			IF pResultCheck <> 0 AND Result = 0 THEN
				Result := pResultCheck;
				codeposition := CONCAT(CONCAT(__POUNAME(),'() / '),__POSITION());
			END_IF;
		END_IF;
		IF pResultCheck = 0 THEN
			count_cycle := 0;
			REPEAT			
				SysFile.SysFileWrite(hFileCheck,ADR(stReSa),TO_UINT(LEN(stReSa)),ADR(pResultCheck));
				count_cycle := count_cycle + 1;
			UNTIL
				pResultCheck = 0 OR count_cycle >= 100 
			END_REPEAT;						
		ELSE
			proError := TRUE;	
			IF Result = 0 THEN
				Result := 16#C7A;
				codeposition := CONCAT(CONCAT(__POUNAME(),'() / '),__POSITION());
			END_IF
		END_IF;  
	END_IF;  
END_IF;
END_METHOD

PROPERTY proFilePathCheckFile : STRING[255];
GET
// FILE Path auf SPS
 proFilePathCheckFile:= CONCAT(  
						CONCAT(  
						CONCAT(                                  
								'$$PlcLogic$$/',  
								'ConfigFiles/Actual/'),  
								stCodeDir),  
								'_Check.txt');
END_GET
END_PROPERTY

METHOD metChild
VAR_INPUT
	itfDataTypeObj  :   ITF_DATATYPE;
END_VAR
IF scState.xGetChild THEN
	IF __QUERYINTERFACE(itfDataTypeObj,itfDataTypeObj) THEN
		IF NOT itfDataTypeObj.proChildAddDone THEN
			usiLastChild := itfDataTypeObj.proparaNr;
			itfDataTypeObj.proChildAddDone := TRUE;
		END_IF;
	END_IF;
END_IF;
END_METHOD

{attribute 'monitoring':='call'}
PROPERTY proLoad : BOOL
GET
proLoad := GVL_Config.xLoad;
END_GET
END_PROPERTY

METHOD FINAL metSaveFile : BOOL
VAR_INPUT  
    itfDataTypeObj  :   ITF_DATATYPE;
END_VAR
VAR
    udiPos  : UDINT;
    stSave  : STRING[172];
	pulPos  : __XWORD;
    dwWrite : DWORD;
	saefty_count	:USINT;
END_VAR
IF hFile <> 0 AND pResult = 0 AND itfDataTypeObj.proParaNr > 0 THEN
    udiPos := LIMIT(1,itfDataTypeObj.proParaNr,255);
   IF udiPos = 1 THEN
        udiPos :=  0;  
        stSave := CONCAT(itfDataTypeObj.proStrPara,'$R'); 
    ELSE
        udiPos := (udiPos * GlobalKonstant.diLineSize) - GlobalKonstant.diLineSize -1;
        stSave := CONCAT('$N',CONCAT(itfDataTypeObj.proStrPara,'$R')); 
	END_IF;
	saefty_count	:= 0;
	REPEAT	
		pResult := SysFile.SysFileSetPos(hFile,0);
		pResult := SysFile.SysFileGetPos(hFile,ADR(pulPos));
		saefty_count := saefty_count + 1;
	UNTIL
		pResult = 0 OR saefty_count >= 10		
	END_REPEAT
	IF pResult <> 0 AND Result = 0 THEN
		Result := pResult;
		codeposition :=   CONCAT(CONCAT(CONCAT(CONCAT(CONCAT(CONCAT(__POUNAME(),'() / '),__POSITION()),' POSW= '),TO_STRING(udiPos)),' POSR='),TO_STRING(pulPos));
		status := SysFile.SysFileGetStatus(hFile);
	END_IF;
	IF pulPos <> udiPos THEN
		saefty_count	:= 0;
		REPEAT
			SysFile.SysFileFlush(hFile);
			pResult := SysFile.SysFileSetPos(hFile,udiPos);
			saefty_count := saefty_count + 1;
		UNTIL
			pResult = 0 OR saefty_count >= 10		
		END_REPEAT
	END_IF;
	IF pResult <> 0 AND Result = 0 THEN
		Result := pResult;
		codeposition :=   CONCAT(CONCAT(CONCAT(CONCAT(CONCAT(CONCAT(__POUNAME(),'() / '),__POSITION()),' POSW= '),TO_STRING(udiPos)),' POSR='),TO_STRING(pulPos));
	END_IF;
    IF hFile <> 0 AND pResult = 0 THEN
		REPEAT 
			pResult := SysFile.SysFileSetPos(hFile,udiPos);
			dwWrite := TO_DWORD(SysFile.SysFileWrite(hFile,ADR(stSave),TO_UDINT(LEN(stSave)),ADR(pResult)));
			SysFile.SysFileFlush(hFile);
			saefty_count := saefty_count + 1;
		UNTIL
			pResult = 0 OR saefty_count >= 10	
		END_REPEAT
		IF pResult <> 0 AND Result = 0 THEN
			Result := pResult;
			codeposition := CONCAT(CONCAT(__POUNAME(),'() / '),__POSITION());
			status := SysFile.SysFileGetStatus(hFile);
		END_IF;
    END_IF;
END_IF;
IF pResult <> 0 THEN
    pResult := pResult;
ELSE
    metSaveFile := NOT TO_BOOL(pResult) AND dwWrite = TO_UDINT(LEN(stSave));
END_IF
scState.xEventSave := TRUE;
END_METHOD

METHOD FINAL metSave : BOOL
VAR_INPUT
    itfDataTypeObj  :   ITF_DATATYPE;
END_VAR
VAR
    uiSafetyCount   :   UINT;
    wPos            :   WORD;
    xSysSemapohre   :   BOOL;
END_VAR
IF proSave OR itfDataTypeObj.proSaveOnChange THEN  
    IF NOT itfDataTypeObj.proIsSaving THEN 
        itfDataTypeObj.proIsSaving := TRUE;
        xSysSemapohre := TRUE;   
    END_IF;
    IF xSysSemapohre THEN
        uiSafetyCount := 0;           
        REPEAT
            pResult := 0; 
            (* File Lesen *)
            IF NOT scState.xIsOpen THEN
                scState.xIsOpen := metOpenFile();
            END_IF;    
            IF scState.xIsOpen THEN
                metSave := metSaveFile(itfDataTypeObj);  
            END_IF;
            uiSafetyCount := uiSafetyCount + 1;
        UNTIL
            metSave = TRUE OR uiSafetyCount = 16#000F
        END_REPEAT
        IF NOT metSave THEN
            THIS^.proError      := TRUE;
            THIS^.proErrorNr    := itfDataTypeObj.proParaNr;
			IF Result = 0 THEN
				Result := 16#C7A;
				codeposition := CONCAT(CONCAT(__POUNAME(),'() / '),__POSITION());
			END_IF
        END_IF  
        xSysSemapohre := FALSE;
        itfDataTypeObj.proIsSaving      := FALSE;
        itfDataTypeObj.proSaveOnChange  := FALSE;		
    END_IF;
END_IF;
END_METHOD

PROPERTY proError : BOOL
GET
proError := xError;
END_GET
SET
xError := proError;
END_SET
END_PROPERTY

{attribute 'monitoring_encoding' := 'UTF-8'}
PROPERTY proFilePath : STRING[255];
GET
// FILE Path auf SPS
proFilePath	     :=      	CONCAT(
							CONCAT(
							CONCAT(                                
									'$$PlcLogic$$/',
									'ConfigFiles/Actual/'),
									stCodeDir),
									'_Config.txt');                                  
								
IF proLoad OR proSave THEN
	proFilePath	    :=      CONCAT(
							CONCAT(
							CONCAT(    
							CONCAT(                            
									'$$PlcLogic$$/',
									'ConfigFiles/'),
									GVL_Config.stBackUp),
									stCodeDir),
									'_Config.txt');  
END_IF;
END_GET
END_PROPERTY

METHOD metCleanUpInit
VAR_INPUT
END_VAR
pResult     		:= fcFileClose(hFile,stCodeDir,'FbConfigFile CleanupIni Z1');
hFile       		:= SysTypes.RTS_INVALID_HANDLE;
pResultCheck		:= fcFileClose(hFileCheck,stCodeDir,'FbConfigFile CleanupIni Z3');
hFileCheck  		:= SysTypes.RTS_INVALID_HANDLE;
fcFileDelete(proFilePathCheckFile);
scState.xInit       := FALSE;
scState.xInitDone	:= TRUE;
iCaseInit   		:= iCaseInit + 1;

IF pResult <> 0 AND Result = 0 THEN
	Result := pResult;
	codeposition := CONCAT(CONCAT(__POUNAME(),'() / '),__POSITION());
END_IF;
IF pResultCheck <> 0 AND Result = 0 THEN
	Result := pResultCheck;
	codeposition := CONCAT(CONCAT(__POUNAME(),'() / '),__POSITION());
END_IF;
END_METHOD

METHOD FINAL metInit : BOOL
VAR_INPUT
    itfDataTypeObj  :   ITF_DATATYPE;
END_VAR
IF scstate.xGetChild THEN
	metChild(itfDataTypeObj);
END_IF;
IF scState.xInit THEN
    IF metCheckNr(itfDataTypeObj,TRUE,FALSE) THEN
        IF NOT metLoadFile(itfDataTypeObj) THEN
            metSaveFile(itfDataTypeObj);
        END_IF;  
        metCheckNr(itfDataTypeObj,FALSE,TRUE);
		metInit := TRUE;
    ELSE    
        proError    := TRUE;
        proErrorNr  := itfDataTypeObj.proParaNr;        
		IF Result = 0 THEN
			Result := 16#C7A;
			codeposition := CONCAT(CONCAT(__POUNAME(),'() / '),__POSITION());
		END_IF
    END_IF;
	IF __QUERYINTERFACE(itfDataTypeObj,itfDataTypeObj) THEN
		IF itfDataTypeObj.proparaNr = usilastChild THEN
			metCleanUpInit();
		END_IF
	END_IF;         
END_IF;
END_METHOD

//FB_Init ist immer implizit verfügbar und wird primär für die Initialisierung verwendet.
//Der Rückgabewert wird nicht ausgewertet. Für gezielte Einflussnahme können Sie
//die Methoden explizit deklarieren und darin mit dem Standard-Initialisierungscode 
//zusätzlichen Code bereitstellen. Sie können den Rückgabewert auswerten.
METHOD FINAL FB_Init: BOOL
VAR_INPUT    
bInitRetains: BOOL; // TRUE: Die Retain-Variablen werden initialisiert (Reset warm / Reset kalt)    
bInCopyCode: BOOL;  // TRUE: Die Instanz wird danach in den Kopiercode kopiert (Online-Change)
END_VAR
hFile   := SysTypes.RTS_INVALID_HANDLE;
hFileCheck  := SysTypes.RTS_INVALID_HANDLE;
END_METHOD

{attribute 'monitoring':='call'}
PROPERTY proSave : BOOL
GET
proSave := GVL_Config.xSave;
END_GET
END_PROPERTY

{attribute 'monitoring':='call'}
PROPERTY proInitDone : BOOL
GET
proInitDone := scState.xInitDone;
END_GET
END_PROPERTY

PROPERTY ProSetInstancePathOnDynCreate : STRING(255)
SET
stCodeDir := ProSetInstancePathOnDynCreate;
metCodeDirCreate();
END_SET
END_PROPERTY

METHOD metCleanUp
VAR_INPUT	
END_VAR
pResult     		:= fcFileClose(hFile,stCodeDir,'FbConfigFile Cleanup Z1');
hFile       		:= SysTypes.RTS_INVALID_HANDLE;
scState.xIsOpen 	:= FALSE;
END_METHOD

METHOD metCheckLastChild
VAR_INPUT  
    itfDataTypeObj  :   ITF_DATATYPE;
END_VAR
IF __QUERYINTERFACE(itfDataTypeObj,itfDataTypeObj) THEN
	IF itfDataTypeObj.proparaNr = usilastChild THEN
		metCleanUp();
	END_IF
END_IF;
END_METHOD

END_FUNCTION_BLOCK

// 30 Program Organization Units/Basis/fbConfigFile
{attribute 'enable_dynamic_creation'}
{attribute 'hide_all_locals'}
{attribute 'reflection'} 
FUNCTION_BLOCK fbConfigFile IMPLEMENTS ITF_CONFIGFILE
VAR_OUTPUT
    xError              :   BOOL;
    uiErrorNr           :   UINT;
	Result              :   RTS_IEC_RESULT;
	codeposition		:	STRING(255);
	status					:	SysFile.SYS_FILE_STATUS;
END_VAR
VAR
    {attribute 'instance-path'} 
    {attribute 'noinit'}     
	{attribute 'monitoring_encoding' := 'UTF-8'}
    stCodeDir               :   STRING[255]; 
    iCaseInit               :   INT                 := 0;
    scState                 :   scStateConfigFile;
    hFile                   :   RTS_IEC_HANDLE;
    pResult                 :   RTS_IEC_RESULT;
    hFileCheck              :   RTS_IEC_HANDLE;
    pResultCheck            :   RTS_IEC_RESULT;    
	usiLastChild			:	USINT;
END_VAR

CASE iCaseInit OF
	0: // Get Last Child
		scState.xGetChild   := TRUE;
		metCodeDirCreate();
		iCaseInit := iCaseInit + 1;
	1: // Init
		scState.xGetChild	:= FALSE;
        scState.xInit       := TRUE;
		
		hFile := fcFileOpen(proFilePath,SysFile.ACCESS_MODE.AM_APPEND_PLUS,pResult);
		IF hFile <> SysTypes.RTS_INVALID_HANDLE THEN
			SysFile.SysFileSetPos(hFile,0);
		END_IF;
		// Check File
		hFileCheck := fcFileOpen(proFilePathCheckFile,SysFile.ACCESS_MODE.AM_WRITE_PLUS,pResultCheck);
		iCaseInit   := iCaseInit + 1;
	2: // Init Done
		;	// Wait on Clean up Init Call
	3: // Check if Save or Load 
		IF (GVL_Config.xSave OR GVL_Config.xLoad) AND_THEN hFile = SysTypes.RTS_INVALID_HANDLE THEN
            scState.xIsOpen := metOpenFile();  
		END_IF;
	ELSE
		iCaseInit   := 0;   
END_CASE;
// Meldung 
IF NOT scState.xEventLoad AND NOT scState.xEventSave AND scState.xEventDetekted THEN
	scState.xEventDetekted := FALSE; 
END_IF;
IF scState.xEventSave THEN
	scState.xEventDetekted := TRUE;
	scState.xEventSave 	   := FALSE;    
END_IF;    
IF scState.xEventLoad THEN
	scState.xEventDetekted := TRUE;
	scState.xEventLoad     := FALSE;    
END_IF; 
IF xError AND_THEN NOT GVL_Config.xError THEN
    GVL_Config.xError 			:= TRUE;
    GVL_Config.stPath			:= stCodeDir;
	GVL_Config.Result			:= Result;
	GVL_Config.codeposition 	:= codeposition;
	GVL_Config.status			:= status;
END_IF;

METHOD FINAL metLoad : BOOL
VAR_INPUT  
    itfDataTypeObj  :   ITF_DATATYPE;
END_VAR
VAR
    uiSafetyCount   :   UINT;
END_VAR
IF proLoad THEN
    REPEAT
        pResult       := 0;
        IF NOT scState.xIsOpen THEN
            scState.xIsOpen := metOpenFile();    
		END_IF
        IF scState.xIsOpen THEN
            metLoad       := metLoadFile(itfDataTypeObj);  
        END_IF;    
            uiSafetyCount := uiSafetyCount + 1;
    UNTIL
        metLoad = TRUE OR uiSafetyCount = 16#FFFF
    END_REPEAT;     
    IF NOT metLoad THEN
        THIS^.proError      := TRUE;
        THIS^.proErrorNr    := itfDataTypeObj.proParaNr;
    END_IF; 
END_IF;
END_METHOD

METHOD metOpenFile : BOOL
VAR_INPUT
END_VAR
hFile   := fcFileOpen(proFilePath,SysFile.ACCESS_MODE.AM_READ_PLUS,pResult);
IF pResult = 0 AND hFile <> SysTypes.RTS_INVALID_HANDLE THEN
    metOpenFile := TRUE;
ELSE
    metOpenFile := FALSE;
END_IF
END_METHOD

PROPERTY proErrorNr : UINT
SET
uiErrorNr := proErrorNr;
END_SET
GET
proErrorNr := uiErrorNr;
END_GET
END_PROPERTY

METHOD PRIVATE FINAL metCodeDirCreate : BOOL
VAR
    uiFor                   :   UINT;
END_VAR
// Instanzpfad des Funktionsbausteinens in Ordnerstrucktur wandeln
FOR uiFor := 0 TO SIZEOF(stCodeDir)-1 DO
    // Punkt . durch Slash / ersetzen
    IF stCodeDir[uiFor] = 46 THEN
        stCodeDir[uiFor] := 47;
    END_IF;            
END_FOR;
END_METHOD

//FB_Exit muss explizit implementiert werden. Wenn es eine Implementierung gibt, dann wird 
//die Methode aufgerufen, bevor die Steuerung den Code der Funktionsbaustein-Instanz entfernt
//(impliziter Aufruf. Der Rückgabewert wird nicht ausgewertet.
METHOD FINAL FB_Exit: BOOL
VAR_INPUT    
    bInCopyCode: BOOL;  // TRUE: Die Exit-Methode wird aufgerufen, um die Instanz zu verlassen, die hinterher kopiert wird Online-Change).  
END_VAR
pResult := SysFile.SysFileClose(hFile);
hFile   := SysTypes.RTS_INVALID_HANDLE;
SysFile.SysFileClose(hFileCheck);
hFileCheck  := SysTypes.RTS_INVALID_HANDLE;
fcFileDelete(proFilePathCheckFile);
END_METHOD

{attribute 'monitoring':='call'}
PROPERTY proSave : BOOL
GET
proSave := GVL_Config.xSave;
END_GET
END_PROPERTY

METHOD FINAL metLoadFile : BOOL
VAR_INPUT  
    itfDataTypeObj  :   ITF_DATATYPE;
END_VAR
VAR
    udiPos  : UDINT;
    stRead  : STRING[170];
    xValid  : BOOL;
END_VAR
IF hFile <> SysTypes.RTS_INVALID_HANDLE AND itfDataTypeObj.proParaNr > 0 THEN
    udiPos := LIMIT(1,itfDataTypeObj.proParaNr,255);
   IF udiPos = 1 THEN
        udiPos :=  udiPos -1;   
    ELSE 
        udiPos := (udiPos * GlobalKonstant.diLineSize) - GlobalKonstant.diLineSize;
	END_IF;
    pResult := SysFile.SysFileSetPos(hFile,udiPos);
END_IF;
IF pResult = 0 AND hFile <> SysTypes.RTS_INVALID_HANDLE THEN
    SysFile.SysFileRead(hFile,ADR(stRead),GlobalKonstant.diStringSize,ADR(pResult));
    stRead[170] := 0;
    IF itfDataTypeObj.proParaNr = TO_UINT(MID(stRead,5,2)) THEN
        itfDataTypeObj.proStrPara := stRead;
        xValid := TRUE;
	END_IF;
END_IF;
metLoadFile := NOT TO_BOOL(pResult) AND xValid;
scState.xEventLoad := TRUE;
END_METHOD

PROPERTY proEventDetekted : BOOL
GET
proEventDetekted := scState.xEventDetekted;
END_GET
END_PROPERTY

METHOD FINAL metCheckNr : BOOL
VAR_INPUT
    itfDataTypeObj  :   ITF_DATATYPE;
    xCheck          :   BOOL;
    xCheckDone      :   BOOL;
END_VAR
VAR
    udiPos  : UDINT;
    stReSa  : STRING[1];
    xValid  : BOOL;
    pulPos  : DWORD;
END_VAR
IF xCheck THEN
    IF pResultCheck = 0 AND itfDataTypeObj.proParaNr > 0 THEN
        udiPos := LIMIT(1,itfDataTypeObj.proParaNr,255)-1;
        pResultCheck := SysFile.SysFileSetPos(hFileCheck,udiPos);
	ELSE
		set_error(CONCAT(CONCAT(__POUNAME(),'() / '),__POSITION()),pResultCheck);
    END_IF;
    IF pResultCheck = 0 THEN
        SysFile.SysFileRead(hFileCheck,ADR(stReSa),1,ADR(pResultCheck));
        IF TO_INT(stReSa) = 1 THEN
            xValid 		:= FALSE; 
			proError 	:= TRUE;
			proErrorNr 	:= itfDataTypeObj.proParaNr;
        ELSE
            xValid := TRUE; 
		END_IF
	ELSE
		proError := TRUE;
		set_error(CONCAT(CONCAT(__POUNAME(),'() / '),__POSITION()),pResultCheck);
    END_IF;
    metCheckNr := NOT TO_BOOL(pResultCheck) AND xValid;
ELSIF xCheckDone THEN
    IF pResultCheck = 0 AND itfDataTypeObj.proParaNr > 0 THEN
            udiPos := LIMIT(1,itfDataTypeObj.proParaNr,255)-1;
            stReSa := TO_STRING(1);
            pResultCheck := SysFile.SysFileGetPos(hFileCheck,ADR(pulPos));
            pResultCheck := SysFile.SysFileSetPos(hFileCheck,udiPos);
            pResultCheck := SysFile.SysFileGetPos(hFileCheck,ADR(pulPos));
    END_IF;
    IF pResultCheck = 0 THEN
        SysFile.SysFileWrite(hFileCheck,ADR(stReSa),TO_UINT(LEN(stReSa)),ADR(pResultCheck));
	ELSE
		set_error(CONCAT(CONCAT(__POUNAME(),'() / '),__POSITION()),pResultCheck);
		proError := TRUE;	
    END_IF;    
END_IF;
END_METHOD

PROPERTY proFilePathCheckFile : STRING[255];
GET
// FILE Path auf SPS
 proFilePathCheckFile:= CONCAT(  
						CONCAT(  
						CONCAT(                                  
								'$$PlcLogic$$/',  
								'ConfigFiles/Actual/'),  
								stCodeDir),  
								'_Check.txt');
END_GET
END_PROPERTY

METHOD metChild
VAR_INPUT
	itfDataTypeObj  :   ITF_DATATYPE;
END_VAR
IF scState.xGetChild THEN
	IF __QUERYINTERFACE(itfDataTypeObj,itfDataTypeObj) THEN
		IF NOT itfDataTypeObj.proChildAddDone THEN
			usiLastChild := itfDataTypeObj.proparaNr;
			itfDataTypeObj.proChildAddDone := TRUE;
		END_IF;
	END_IF;
END_IF;
END_METHOD

PROPERTY proError : BOOL
GET
proError := xError;
END_GET
SET
xError := proError;
END_SET
END_PROPERTY

{attribute 'monitoring':='call'}
PROPERTY proLoad : BOOL
GET
proLoad := GVL_Config.xLoad;
END_GET
END_PROPERTY

METHOD FINAL metSaveFile : BOOL
VAR_INPUT  
    itfDataTypeObj  :   ITF_DATATYPE;
END_VAR
VAR
    udiPos  : UDINT;
    stSave  : STRING[172];
	pulPos  : DWORD;
    dwWrite : DWORD;
END_VAR
IF hFile <> SysTypes.RTS_INVALID_HANDLE AND pResult = 0 AND itfDataTypeObj.proParaNr > 0 THEN
    udiPos := LIMIT(1,itfDataTypeObj.proParaNr,255);
   IF udiPos = 1 THEN
        udiPos :=  udiPos -1;  
        stSave := CONCAT(itfDataTypeObj.proStrPara,'$R'); 
    ELSE
        udiPos := (udiPos * GlobalKonstant.diLineSize) - GlobalKonstant.diLineSize - 1;
        stSave := CONCAT('$N',CONCAT(itfDataTypeObj.proStrPara,'$R')); 
	END_IF;
        pResult := SysFile.SysFileGetPos(hFile,ADR(pulPos));
        pResult := SysFile.SysFileSetPos(hFile,udiPos);
        pResult := SysFile.SysFileGetPos(hFile,ADR(pulPos));
    IF hFile <> 0 AND pResult = 0 THEN
        dwWrite := TO_DWORD(SysFile.SysFileWrite(hFile,ADR(stSave),TO_UDINT(LEN(stSave)),ADR(pResult)));
	ELSE
		set_error(CONCAT(CONCAT(__POUNAME(),'() / '),__POSITION()),pResult);
    END_IF;
END_IF;
IF pResult <> 0 THEN
	set_error(CONCAT(CONCAT(__POUNAME(),'() / '),__POSITION()),pResult);
ELSE
    metSaveFile := NOT TO_BOOL(pResult) AND dwWrite = TO_UDINT(LEN(stSave));
END_IF
scState.xEventSave := TRUE;
END_METHOD

METHOD FINAL metSave : BOOL
VAR_INPUT
    itfDataTypeObj  :   ITF_DATATYPE;
END_VAR
VAR
    uiSafetyCount   :   UINT;
    wPos            :   WORD;
    xSysSemapohre   :   BOOL;
END_VAR
IF NOT xError THEN
	IF proSave OR itfDataTypeObj.proSaveOnChange THEN  
		IF NOT itfDataTypeObj.proIsSaving THEN 
			itfDataTypeObj.proIsSaving := TRUE;
			xSysSemapohre := TRUE;   
		END_IF;
		IF xSysSemapohre THEN
			uiSafetyCount := 0;           
			REPEAT
				pResult := 0; 
				(* File Lesen *)
				IF NOT scState.xIsOpen THEN
					scState.xIsOpen := metOpenFile();
				END_IF;    
				IF scState.xIsOpen THEN
					metSave := metSaveFile(itfDataTypeObj);  
				END_IF;
				uiSafetyCount := uiSafetyCount + 1;
				IF NOT metSave THEN
					wPos := 16#EEEE;    
				END_IF
			UNTIL
				metSave = TRUE OR uiSafetyCount = 16#FFFF
			END_REPEAT
			IF NOT metSave THEN
				THIS^.proError      := TRUE;
				THIS^.proErrorNr    := itfDataTypeObj.proParaNr;
			END_IF  
			xSysSemapohre := FALSE;
			itfDataTypeObj.proIsSaving      := FALSE;
			itfDataTypeObj.proSaveOnChange  := FALSE;		
		END_IF;
	END_IF;
END_IF;
END_METHOD

{attribute 'monitoring':='call'}
PROPERTY proInitDone : BOOL
GET
proInitDone := scState.xInitDone;
END_GET
END_PROPERTY

{attribute 'monitoring_encoding' := 'UTF-8'}
PROPERTY proFilePath : STRING[255];
GET
// FILE Path auf SPS
proFilePath     :=      	CONCAT(
							CONCAT(
							CONCAT(                                
									'$$PlcLogic$$/',
									'ConfigFiles/Actual/'),
									stCodeDir),
									'_Config.txt');                                  
								
IF proLoad OR proSave THEN
	proFilePath     :=      CONCAT(
							CONCAT(
							CONCAT(    
							CONCAT(                            
									'$$PlcLogic$$/',
									'ConfigFiles/'),
									GVL_Config.stBackUp),
									stCodeDir),
									'_Config.txt');  
END_IF;
END_GET
END_PROPERTY

METHOD metCleanUpInit
VAR_INPUT
END_VAR
pResult     		:= fcFileClose(hFile,stCodeDir,'FbConfigFile CleanupIni Z1');
hFile       		:= SysTypes.RTS_INVALID_HANDLE;
pResultCheck		:= fcFileClose(hFileCheck,stCodeDir,'FbConfigFile CleanupIni Z3');
hFileCheck  		:= SysTypes.RTS_INVALID_HANDLE;
fcFileDelete(proFilePathCheckFile);
scState.xInit       := FALSE;
scState.xInitDone	:= TRUE;
iCaseInit   		:= iCaseInit + 1;
END_METHOD

METHOD FINAL metInit : BOOL
VAR_INPUT
    itfDataTypeObj  :   ITF_DATATYPE;
END_VAR
IF scstate.xGetChild THEN
	metChild(itfDataTypeObj);
END_IF;
IF scState.xInit THEN
    IF metCheckNr(itfDataTypeObj,TRUE,FALSE) THEN
        IF NOT metLoadFile(itfDataTypeObj) THEN
            metSaveFile(itfDataTypeObj);
        END_IF;  
        metCheckNr(itfDataTypeObj,FALSE,TRUE);
		metInit := TRUE;
    ELSE    
        proError    := TRUE;
        proErrorNr  := itfDataTypeObj.proParaNr;        
    END_IF;
	IF __QUERYINTERFACE(itfDataTypeObj,itfDataTypeObj) THEN
		IF itfDataTypeObj.proparaNr = usilastChild THEN
			metCleanUpInit();
		END_IF
	END_IF;         
END_IF;
END_METHOD

//FB_Init ist immer implizit verfügbar und wird primär für die Initialisierung verwendet.
//Der Rückgabewert wird nicht ausgewertet. Für gezielte Einflussnahme können Sie
//die Methoden explizit deklarieren und darin mit dem Standard-Initialisierungscode 
//zusätzlichen Code bereitstellen. Sie können den Rückgabewert auswerten.
METHOD FINAL FB_Init: BOOL
VAR_INPUT    
bInitRetains: BOOL; // TRUE: Die Retain-Variablen werden initialisiert (Reset warm / Reset kalt)    
bInCopyCode: BOOL;  // TRUE: Die Instanz wird danach in den Kopiercode kopiert (Online-Change)
END_VAR
hFile   := SysTypes.RTS_INVALID_HANDLE;
hFileCheck  := SysTypes.RTS_INVALID_HANDLE;
END_METHOD

PROPERTY ProSetInstancePathOnDynCreate : STRING(255)
SET
stCodeDir := ProSetInstancePathOnDynCreate;
metCodeDirCreate();
END_SET
END_PROPERTY

METHOD metCleanUp
VAR_INPUT	
END_VAR
pResult     		:= fcFileClose(hFile,stCodeDir,'FbConfigFile Cleanup Z1');
hFile       		:= SysTypes.RTS_INVALID_HANDLE;
scState.xIsOpen 	:= FALSE;
END_METHOD

METHOD metCheckLastChild
VAR_INPUT  
    itfDataTypeObj  :   ITF_DATATYPE;
END_VAR
IF __QUERYINTERFACE(itfDataTypeObj,itfDataTypeObj) THEN
	IF itfDataTypeObj.proparaNr = usilastChild THEN
		metCleanUp();
	END_IF
END_IF;
END_METHOD

METHOD set_error
VAR_INPUT
	_codeposition : STRING(255);
	_ResultIn	  : RTS_IEC_RESULT;
END_VAR
IF Result = 0 THEN
	Result := _ResultIn;
	codeposition := _codeposition;
END_IF;
END_METHOD

END_FUNCTION_BLOCK

// 30 Program Organization Units/40 Byte String/fbSTRING40
FUNCTION_BLOCK fbSTRING40 EXTENDS fbDataType IMPLEMENTS ITF_STRING40
VAR_INPUT CONSTANT
	{attribute 'monitoring_encoding' := 'UTF-8'}
    _WertInit      :   STRING[40];  
END_VAR
VAR
	{attribute 'monitoring_encoding' := 'UTF-8'}
    stValue          :   STRING[40]; 
    {attribute 'hide'}
	{attribute 'monitoring_encoding' := 'UTF-8'}
    stValueOld       :   STRING[40]; 
END_VAR

(* Call Supper Objekt *)
IF itfConfigFb <> 0 THEN
    SUPER^();
END_IF;

{attribute 'hide'}
{attribute 'monitoring':='call'}
{attribute 'monitoring_encoding' := 'UTF-8'}
PROPERTY proStrPara : STRING(129)
// {attribute 'hide'}
GET
proStrPara :=   CONCAT(                    
                CONCAT( 
                CONCAT(
                CONCAT(                 
                CONCAT(                     
                CONCAT( fcfillStr(CONCAT('P',TO_STRING(SUPER^._usiParaNr)),6)       ,
                        ';'                                                         ),
                        fcfillStr(TO_STRING(stValue),GlobalKonstant.usiFeldLeng)    ),
                        ';'                                                         ),
                        fcfillStr('',GlobalKonstant.usiFeldLeng)                    ),
                        ';'                                                         ),
                        fcfillStr('',GlobalKonstant.usiFeldLeng)                    );
END_GET
SET
proValue  := fcGetValue(proStrPara);
END_SET
END_PROPERTY

METHOD metNewValueNoSave : BOOL
VAR_INPUT
    newValueNoSave   :   STRING[40];
END_VAR
proValue := newValueNoSave;
scState.xUpdateOldValueNoSave := TRUE;
metNewValueNoSave := TRUE;
END_METHOD

{attribute 'hide'}
METHOD metInit : BOOL
proValue  := _WertInit;
END_METHOD

{attribute 'monitoring_encoding' := 'UTF-8'}
PROPERTY proShowValue : STRING[40]
GET
proShowValue := stValue;
END_GET
END_PROPERTY

{attribute 'monitoring':='call'}
{attribute 'monitoring_encoding' := 'UTF-8'}
PROPERTY proValue : STRING[40]
SET
stValue := proValue;
(* Hack da Virtual Keyboard kein ° Zeichen hat *)
IF FIND(stValue,'§C') > 0 THEN
    stValue := REPLACE(stValue,'°',1,FIND(stValue,'§C'));
END_IF;
stValue[40] := 0;
END_SET
GET
stValue[40] := 0;
proValue := stValue;
END_GET
END_PROPERTY

METHOD metNewValue : BOOL
VAR_INPUT
    newValue   :   STRING[40];
END_VAR
proValue := newValue;
metNewValue := TRUE;
END_METHOD

{attribute 'hide'}
METHOD metCheckState : BOOL
(* Search Change & Save Old Values *)
IF stValue <> stValueOld OR scState.xUpdateOldValueNoSave THEN
    (* Prüfen ob die Werte bei änderung gespeichert werden sollen *)
    IF scState.xUpdateOldValueNoSave THEN
        scState.xUpdateOldValueNoSave := FALSE;
    ELSE
        proSaveOnChange 	:= TRUE;
	END_IF
	(*State Changed*) 
	scState.xStateChanged 	:= TRUE;   
    proValue 				:= stValue;
    stValueOld 				:= proValue;
ELSE
	(*State Changed*) 
	scState.xStateChanged 	:= FALSE;    
END_IF;
END_METHOD

END_FUNCTION_BLOCK

// 40 Visualizations/32 Bit/DWORD/DWORD DEZ/visDWORD_QUERRY_DEZ
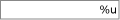
VISUALIZATION visDWORD_QUERRY_DEZ  // 120x20
VAR_INPUT
    visfbDWORDIn :   ITF_DWORD;	
END_VAR
    Frame (0,0 120x20), invisible if: NOT __QUERYINTERFACE(visfbDWORDIn,visfbDWORDIn)
        shows visDWORD_ITF_DEZ(visfbDWORD := visfbDWORDIn)
END_VISUALIZATION

// 40 Visualizations/1 Bit/visBOOL
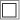
VISUALIZATION visBOOL  // 20x20
VAR_INPUT
    visfbBOOLIn  : ITF_DATATYPE;
END_VAR
VAR    
    visfbBOOL    : ITF_BOOL;    	
END_VAR
    Frame (0,0 20x20), invisible if: NOT __QUERYINTERFACE(visfbBOOLIn,visfbBOOL)
        shows visBOOL_QUERRY(visfbBOOLIn := visfbBOOL)
END_VISUALIZATION

// 40 Visualizations/32 Bit/UDINT/visUDINT
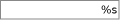
VISUALIZATION visUDINT  // 120x20
VAR_INPUT
    visfbUDINTIn :   ITF_DATATYPE;	
END_VAR
VAR
    visfbUDINT   :   ITF_UDINT;	
END_VAR
VAR_INPUT 
    stPhysikalischeEinheit  : STRING[5];
END_VAR
    Frame (0,0 120x20), invisible if: NOT __QUERYINTERFACE(visfbUDINTIn,visfbUDINT)
        shows visUDINT_QUERRY(visfbUDINTIn := visfbUDINT, stPhysikalischeEinheit := stPhysikalischeEinheit)
END_VISUALIZATION

// 40 Visualizations/32 Bit/TIME/visTIME
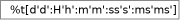
VISUALIZATION visTIME  // 180x20
VAR_INPUT   
    visfbTIMEIn :   ITF_DATATYPE;	
END_VAR
VAR  
    visfbTIME   :   ITF_TIME;	
END_VAR
    Frame (0,0 180x20), invisible if: NOT __QUERYINTERFACE(visfbTIMEIn,visfbTIME)
        shows visTIME_QUERRY(visfbTIMEIn := visfbTIME)
END_VISUALIZATION

// 40 Visualizations/32 Bit/REAL/visREAL_QUERRY
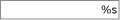
VISUALIZATION visREAL_QUERRY  // 120x20
VAR_INPUT    
    visfbREALIn :   ITF_REAL;	
END_VAR
VAR_INPUT 
    stPhysikalischeEinheit  : STRING[5];
END_VAR
    Frame (0,0 120x20), invisible if: NOT __QUERYINTERFACE(visfbREALIn,visfbREALIn)
        shows visREAL_ITF(visfbREAL := visfbREALIn, stPhysikalischeEinheit := stPhysikalischeEinheit)
END_VISUALIZATION

// 40 Visualizations/1 Bit/visBOOL_ITF
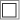
VISUALIZATION visBOOL_ITF  // 20x20
VAR_INPUT
    visfbBOOL    : ITF_BOOL;    	
END_VAR
    Checkbox (0,0 20x20), variable: visfbBOOL.proValue
END_VISUALIZATION

// 40 Visualizations/ENUMERATION/32 Bit/visENUMERATION_DINT_QUERRY
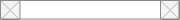
VISUALIZATION visENUMERATION_DINT_QUERRY  // 180x20
VAR_INPUT
    visfbDINT   :   ITF_DINT;	
END_VAR
    Frame (0,0 180x20), invisible if: NOT __QUERYINTERFACE(visfbDINT,visfbDINT)
        shows visENUMERATION_DINT(visfbDINT := visfbDINT)
END_VISUALIZATION

// 40 Visualizations/16 Bit/WORD/WORD HEX/visWORD_HEX
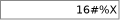
VISUALIZATION visWORD_HEX  // 120x20
VAR_INPUT
    visfbWORDIn :   ITF_DATATYPE;	
END_VAR
VAR
    visfbWORD   :   ITF_WORD;	
END_VAR
    Frame (0,0 120x20), invisible if: NOT __QUERYINTERFACE(visfbWORDIn,visfbWORD)
        shows visWORD_QUERRY_HEX(visfbWORDIn := visfbWORD)
END_VISUALIZATION

// 40 Visualizations/64 Bit/LTIME/visLTIME_ITF
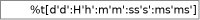
VISUALIZATION visLTIME_ITF  // 200x20
VAR_INPUT
    visfbLTIME   :   ITF_LTIME;	
END_VAR
    Textfield (0,0 200x20), "%t[d'd':H'h':m'm':ss's':ms'ms']", text variable: visfbLTIME.proValue
        OnMouseClick: write the text variable via InputWithLimits, min TO_ULINT(visfbLTIME.proMin), max TO_ULINT(visfbLTIME.proMax), title 'T#'
END_VISUALIZATION

// 40 Visualizations/32 Bit/REAL/visREAL
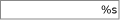
VISUALIZATION visREAL  // 120x20
VAR_INPUT
    visfbREALIn :   ITF_DATATYPE;	
END_VAR
VAR
    visfbREAL   :   ITF_REAL;	
END_VAR
VAR_INPUT 
    stPhysikalischeEinheit  : STRING[5];
END_VAR
    Frame (0,0 120x20), invisible if: NOT __QUERYINTERFACE(visfbREALIn,visfbREAL)
        shows visREAL_QUERRY(visfbREALIn := visfbREAL, stPhysikalischeEinheit := stPhysikalischeEinheit)
END_VISUALIZATION

// 40 Visualizations/32 Bit/DATE AND TIME/visDATE_AND_TIME_ITF
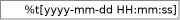
VISUALIZATION visDATE_AND_TIME_ITF  // 180x20
VAR_INPUT
    visfbDATE_AND_TIMEIn   :   ITF_DATE_AND_TIME;	
END_VAR
    Textfield (0,0 180x20), "%t[yyyy-mm-dd HH:mm:ss]", text variable: visfbDATE_AND_TIMEIn.proValue
        OnMouseClick: write the text variable via InputWithLimits, min TO_UDINT(visfbDATE_AND_TIMEIn.proMin), max TO_UDINT(visfbDATE_AND_TIMEIn.proMax), title 'T#'
END_VISUALIZATION

// 40 Visualizations/16 Bit/INT/visINT
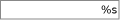
VISUALIZATION visINT  // 120x20
VAR_INPUT
    visfbINTIn :   ITF_DATATYPE;	
END_VAR
VAR
    visfbINT   :   ITF_INT;	
END_VAR
VAR_INPUT 
    stPhysikalischeEinheit  : STRING[5];
END_VAR
    Frame (0,0 120x20), invisible if: NOT __QUERYINTERFACE(visfbINTIn,visfbINT)
        shows visINT_QUERRY(visfbINTIn := visfbINT, stPhysikalischeEinheit := stPhysikalischeEinheit)
END_VISUALIZATION

// 40 Visualizations/32 Bit/UDINT/visUDINT_QUERRY
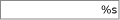
VISUALIZATION visUDINT_QUERRY  // 120x20
VAR_INPUT
    visfbUDINTIn :   ITF_UDINT;	
END_VAR
VAR_INPUT 
    stPhysikalischeEinheit  : STRING[5];
END_VAR
    Frame (0,0 120x20), invisible if: NOT __QUERYINTERFACE(visfbUDINTIn,visfbUDINTIn)
        shows visUDINT_ITF(visfbUDINT := visfbUDINTIn, stPhysikalischeEinheit := stPhysikalischeEinheit)
END_VISUALIZATION

// 40 Visualizations/8 Bit/SINT/visSINT_QUERRY
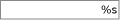
VISUALIZATION visSINT_QUERRY  // 120x20
VAR_INPUT
    visfbSINTIn :   ITF_SINT;	
END_VAR
VAR_INPUT 
    stPhysikalischeEinheit  : STRING[5];
END_VAR
    Frame (0,0 120x20), invisible if: NOT __QUERYINTERFACE(visfbSINTIn,visfbSINTIn)
        shows visSINT_ITF(visfbSINT := visfbSINTIn, stPhysikalischeEinheit := stPhysikalischeEinheit)
END_VISUALIZATION

// 40 Visualizations/16 Bit/WORD/WORD DEZ/visWORD_ITF_DEZ
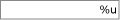
VISUALIZATION visWORD_ITF_DEZ  // 120x20
VAR_INPUT
    visfbWORD   :   ITF_WORD;	
END_VAR
    Textfield (0,0 120x20), "%u", text variable: visfbWORD.proValue
        OnMouseClick: write the text variable via InputWithLimits, min visfbWORD.proMin, max visfbWORD.proMax
END_VISUALIZATION

// 40 Visualizations/32 Bit/TOD/visTOD_ITF
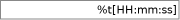
VISUALIZATION visTOD_ITF  // 180x20
VAR_INPUT
    visfbTODIn   :   ITF_TOD;	
END_VAR
    Textfield (0,0 180x20), "%t[HH:mm:ss]", text variable: visfbTODIn.proValue
        OnMouseClick: write the text variable via InputWithLimits, min TO_UDINT(visfbTODIn.proMin), max TO_UDINT(visfbTODIn.proMax), title 'Tod#'
END_VISUALIZATION

// 40 Visualizations/16 Bit/INT/visINT_ITF
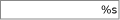
VISUALIZATION visINT_ITF  // 120x20
VAR_INPUT
    visfbINT   :   ITF_INT;	
END_VAR
VAR_INPUT 
    stPhysikalischeEinheit  : STRING[5];
END_VAR
    Textfield (0,0 120x20), "%s", text variable: CONCAT(TO_STRING(visfbINT.proValue),stPhysikalischeEinheit)
        OnMouseClick: write visfbINT.proValue via InputWithLimits, min visfbINT.proMin, max visfbINT.proMax
END_VISUALIZATION

// 40 Visualizations/8 Bit/USINT/visUSINT_QUERRY
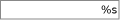
VISUALIZATION visUSINT_QUERRY  // 120x20
VAR_INPUT
    visfbUSINTIn :   ITF_USINT;	
END_VAR
VAR_INPUT 
    stPhysikalischeEinheit  : STRING[5];
END_VAR
    Frame (0,0 120x20), invisible if: NOT __QUERYINTERFACE(visfbUSINTIn,visfbUSINTIn)
        shows visUSINT_ITF(visfbUSINT := visfbUSINTIn, stPhysikalischeEinheit := stPhysikalischeEinheit)
END_VISUALIZATION

// 40 Visualizations/8 Bit/USINT/visUSINT_ITF
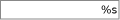
VISUALIZATION visUSINT_ITF  // 120x20
VAR_INPUT
    visfbUSINT   :   ITF_USINT;	
END_VAR
VAR_INPUT 
    stPhysikalischeEinheit  : STRING[5];
END_VAR
    Textfield (0,0 120x20), "%s", text variable: CONCAT(TO_STRING(visfbUSINT.proValue),stPhysikalischeEinheit)
        OnMouseClick: write visfbUSINT.proValue via InputWithLimits, min visfbUSINT.proMin, max visfbUSINT.proMax
END_VISUALIZATION

// 40 Visualizations/40 Byte String/visSTRING40_QUERRY
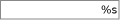
VISUALIZATION visSTRING40_QUERRY  // 120x20
VAR_INPUT
    visfbSTRING40In :   ITF_STRING40;	
END_VAR
    Frame (0,0 120x20), invisible if: NOT __QUERYINTERFACE(visfbSTRING40In,visfbSTRING40In)
        shows visSTRING40_ITF(visfbSTRING40In := visfbSTRING40In)
END_VISUALIZATION

// 40 Visualizations/16 Bit/WORD/WORD DEZ/visWORD_QUERRY_DEZ
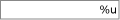
VISUALIZATION visWORD_QUERRY_DEZ  // 120x20
VAR_INPUT
    visfbWORDIn :   ITF_WORD;	
END_VAR
    Frame (0,0 120x20), invisible if: NOT __QUERYINTERFACE(visfbWORDIn,visfbWORDIn)
        shows visWORD_ITF_DEZ(visfbWORD := visfbWORDIn)
END_VISUALIZATION

// 40 Visualizations/40 Byte String/visSTRING40
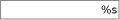
VISUALIZATION visSTRING40  // 120x20
VAR_INPUT
    visfbSTRING40In :   ITF_DATATYPE;	
END_VAR
VAR
    visfbSTRING40   :   ITF_STRING40;	
END_VAR
    Frame (0,0 120x20), invisible if: NOT __QUERYINTERFACE(visfbSTRING40In,visfbSTRING40)
        shows visSTRING40_QUERRY(visfbSTRING40In := visfbSTRING40)
END_VISUALIZATION

// 40 Visualizations/64 Bit/LTIME/visLTIME
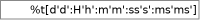
VISUALIZATION visLTIME  // 200x20
VAR_INPUT   
    visfbLTIMEIn :   ITF_DATATYPE;	
END_VAR
VAR  
    visfbLTIME   :   ITF_LTIME;	
END_VAR
    Frame (0,0 200x20), invisible if: NOT __QUERYINTERFACE(visfbLTIMEIn,visfbLTIME)
        shows visLTIME_QUERRY(visfbLTIMEIn := visfbLTIME)
END_VISUALIZATION

// 40 Visualizations/16 Bit/WORD/WORD DEZ/visWORD_DEZ
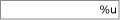
VISUALIZATION visWORD_DEZ  // 120x20
VAR_INPUT
    visfbWORDIn :   ITF_DATATYPE;	
END_VAR
VAR
    visfbWORD   :   ITF_WORD;	
END_VAR
    Frame (0,0 120x20), invisible if: NOT __QUERYINTERFACE(visfbWORDIn,visfbWORD)
        shows visWORD_QUERRY_DEZ(visfbWORDIn := visfbWORD)
END_VISUALIZATION

// 40 Visualizations/Show Data/visSHOWDATA_QUERRY
